(* IEC 61131-3 sources: taksa-factory-simulator/sample_programs, 16 files *)

(* ---- CNCMachiningPLC10.st ---- *)
PROGRAM PLC10_CNC

VAR
    cycle_time : REAL := 120.0;
    throughput : REAL := 30.0;

    dimension_ok : BOOL := TRUE;
    surface_finish : REAL := 0.95;

    tool_break_alarm : BOOL := FALSE;

    spindle_energy : REAL := 50.0;

    machine_idle : REAL := 0.0;

    spindle_load : REAL := 70.0;
    tool_life : REAL := 100.0;

    rand : REAL;
    tick : DINT;
END_VAR

VAR_EXTERNAL
    reg_cycle_time_x10 : UINT;
    reg_throughput_x10 : UINT;
    reg_dimension_ok : UINT;
    reg_surface_finish_x1000 : UINT;
    reg_tool_break_alarm : UINT;
    reg_spindle_energy_x10 : UINT;
    reg_machine_idle_x10 : UINT;
    reg_spindle_load_x10 : UINT;
    reg_tool_life_x10 : UINT;
END_VAR

rand := DINT_TO_REAL((tick * 41) MOD 100) / 100.0;
tick := tick + 1;

cycle_time := 100.0 + (rand * 40.0);
throughput := 3600.0 / cycle_time;

spindle_load := 60.0 + (rand * 30.0);

IF rand < 0.01 THEN
    tool_break_alarm := TRUE;
    dimension_ok := FALSE;
END_IF;

tool_life := tool_life - 0.001;

spindle_energy := spindle_load * 0.8;

(* Export live values to Modbus holding registers %MW0.. *)
reg_cycle_time_x10 := REAL_TO_UINT(cycle_time * 10.0);
reg_throughput_x10 := REAL_TO_UINT(throughput * 10.0);
IF dimension_ok THEN
    reg_dimension_ok := 1;
ELSE
    reg_dimension_ok := 0;
END_IF;
reg_surface_finish_x1000 := REAL_TO_UINT(surface_finish * 1000.0);
IF tool_break_alarm THEN
    reg_tool_break_alarm := 1;
ELSE
    reg_tool_break_alarm := 0;
END_IF;
reg_spindle_energy_x10 := REAL_TO_UINT(spindle_energy * 10.0);
reg_machine_idle_x10 := REAL_TO_UINT(machine_idle * 10.0);
reg_spindle_load_x10 := REAL_TO_UINT(spindle_load * 10.0);
reg_tool_life_x10 := REAL_TO_UINT(tool_life * 10.0);

END_PROGRAM

CONFIGURATION Config0
  RESOURCE Res0 ON PLC
    VAR_GLOBAL
      reg_cycle_time_x10 AT %MW0 : UINT;
      reg_throughput_x10 AT %MW1 : UINT;
      reg_dimension_ok AT %MW2 : UINT;
      reg_surface_finish_x1000 AT %MW3 : UINT;
      reg_tool_break_alarm AT %MW4 : UINT;
      reg_spindle_energy_x10 AT %MW5 : UINT;
      reg_machine_idle_x10 AT %MW6 : UINT;
      reg_spindle_load_x10 AT %MW7 : UINT;
      reg_tool_life_x10 AT %MW8 : UINT;
    END_VAR

    TASK Main(INTERVAL := T#20ms, PRIORITY := 0);
    PROGRAM Inst0 WITH Main : PLC10_CNC;
  END_RESOURCE
END_CONFIGURATION

(* ---- CNCMachiningPLC8.st ---- *)
PROGRAM PLC8_CNC

VAR
    cycle_time : REAL := 120.0;
    throughput : REAL := 30.0;

    dimension_ok : BOOL := TRUE;
    surface_finish : REAL := 0.95;

    tool_break_alarm : BOOL := FALSE;

    spindle_energy : REAL := 50.0;

    machine_idle : REAL := 0.0;

    spindle_load : REAL := 70.0;
    tool_life : REAL := 100.0;

    rand : REAL;
    tick : DINT;
END_VAR

VAR_EXTERNAL
    reg_cycle_time_x10 : UINT;
    reg_throughput_x10 : UINT;
    reg_dimension_ok : UINT;
    reg_surface_finish_x1000 : UINT;
    reg_tool_break_alarm : UINT;
    reg_spindle_energy_x10 : UINT;
    reg_machine_idle_x10 : UINT;
    reg_spindle_load_x10 : UINT;
    reg_tool_life_x10 : UINT;
END_VAR

rand := DINT_TO_REAL((tick * 41) MOD 100) / 100.0;
tick := tick + 1;

cycle_time := 100.0 + (rand * 40.0);
throughput := 3600.0 / cycle_time;

spindle_load := 60.0 + (rand * 30.0);

IF rand < 0.01 THEN
    tool_break_alarm := TRUE;
    dimension_ok := FALSE;
END_IF;

tool_life := tool_life - 0.001;

spindle_energy := spindle_load * 0.8;

(* Export live values to Modbus holding registers %MW0.. *)
reg_cycle_time_x10 := REAL_TO_UINT(cycle_time * 10.0);
reg_throughput_x10 := REAL_TO_UINT(throughput * 10.0);
IF dimension_ok THEN
    reg_dimension_ok := 1;
ELSE
    reg_dimension_ok := 0;
END_IF;
reg_surface_finish_x1000 := REAL_TO_UINT(surface_finish * 1000.0);
IF tool_break_alarm THEN
    reg_tool_break_alarm := 1;
ELSE
    reg_tool_break_alarm := 0;
END_IF;
reg_spindle_energy_x10 := REAL_TO_UINT(spindle_energy * 10.0);
reg_machine_idle_x10 := REAL_TO_UINT(machine_idle * 10.0);
reg_spindle_load_x10 := REAL_TO_UINT(spindle_load * 10.0);
reg_tool_life_x10 := REAL_TO_UINT(tool_life * 10.0);

END_PROGRAM

CONFIGURATION Config0
  RESOURCE Res0 ON PLC
    VAR_GLOBAL
      reg_cycle_time_x10 AT %MW0 : UINT;
      reg_throughput_x10 AT %MW1 : UINT;
      reg_dimension_ok AT %MW2 : UINT;
      reg_surface_finish_x1000 AT %MW3 : UINT;
      reg_tool_break_alarm AT %MW4 : UINT;
      reg_spindle_energy_x10 AT %MW5 : UINT;
      reg_machine_idle_x10 AT %MW6 : UINT;
      reg_spindle_load_x10 AT %MW7 : UINT;
      reg_tool_life_x10 AT %MW8 : UINT;
    END_VAR

    TASK Main(INTERVAL := T#20ms, PRIORITY := 0);
    PROGRAM Inst0 WITH Main : PLC8_CNC;
  END_RESOURCE
END_CONFIGURATION

(* ---- CNCMachiningPLC9.st ---- *)
PROGRAM PLC9_CNC

VAR
    cycle_time : REAL := 120.0;
    throughput : REAL := 30.0;

    dimension_ok : BOOL := TRUE;
    surface_finish : REAL := 0.95;

    tool_break_alarm : BOOL := FALSE;

    spindle_energy : REAL := 50.0;

    machine_idle : REAL := 0.0;

    spindle_load : REAL := 70.0;
    tool_life : REAL := 100.0;

    rand : REAL;
    tick : DINT;
END_VAR

VAR_EXTERNAL
    reg_cycle_time_x10 : UINT;
    reg_throughput_x10 : UINT;
    reg_dimension_ok : UINT;
    reg_surface_finish_x1000 : UINT;
    reg_tool_break_alarm : UINT;
    reg_spindle_energy_x10 : UINT;
    reg_machine_idle_x10 : UINT;
    reg_spindle_load_x10 : UINT;
    reg_tool_life_x10 : UINT;
END_VAR

rand := DINT_TO_REAL((tick * 41) MOD 100) / 100.0;
tick := tick + 1;

cycle_time := 100.0 + (rand * 40.0);
throughput := 3600.0 / cycle_time;

spindle_load := 60.0 + (rand * 30.0);

IF rand < 0.01 THEN
    tool_break_alarm := TRUE;
    dimension_ok := FALSE;
END_IF;

tool_life := tool_life - 0.001;

spindle_energy := spindle_load * 0.8;

(* Export live values to Modbus holding registers %MW0.. *)
reg_cycle_time_x10 := REAL_TO_UINT(cycle_time * 10.0);
reg_throughput_x10 := REAL_TO_UINT(throughput * 10.0);
IF dimension_ok THEN
    reg_dimension_ok := 1;
ELSE
    reg_dimension_ok := 0;
END_IF;
reg_surface_finish_x1000 := REAL_TO_UINT(surface_finish * 1000.0);
IF tool_break_alarm THEN
    reg_tool_break_alarm := 1;
ELSE
    reg_tool_break_alarm := 0;
END_IF;
reg_spindle_energy_x10 := REAL_TO_UINT(spindle_energy * 10.0);
reg_machine_idle_x10 := REAL_TO_UINT(machine_idle * 10.0);
reg_spindle_load_x10 := REAL_TO_UINT(spindle_load * 10.0);
reg_tool_life_x10 := REAL_TO_UINT(tool_life * 10.0);

END_PROGRAM

CONFIGURATION Config0
  RESOURCE Res0 ON PLC
    VAR_GLOBAL
      reg_cycle_time_x10 AT %MW0 : UINT;
      reg_throughput_x10 AT %MW1 : UINT;
      reg_dimension_ok AT %MW2 : UINT;
      reg_surface_finish_x1000 AT %MW3 : UINT;
      reg_tool_break_alarm AT %MW4 : UINT;
      reg_spindle_energy_x10 AT %MW5 : UINT;
      reg_machine_idle_x10 AT %MW6 : UINT;
      reg_spindle_load_x10 AT %MW7 : UINT;
      reg_tool_life_x10 AT %MW8 : UINT;
    END_VAR

    TASK Main(INTERVAL := T#20ms, PRIORITY := 0);
    PROGRAM Inst0 WITH Main : PLC9_CNC;
  END_RESOURCE
END_CONFIGURATION

(* ---- Cooling.st ---- *)
PROGRAM PLC5_COOLING

VAR
    cooling_time : REAL := 120.0;

    cooling_uniformity : REAL := 0.95;

    temp_alarm : BOOL := FALSE;

    water_usage : REAL := 50.0;

    blockage_time : REAL := 0.0;

    pump_health : REAL := 100.0;

    rand : REAL;
    tick : DINT;
END_VAR

VAR_EXTERNAL
    reg_cooling_time_x10 : UINT;
    reg_cooling_uniformity_x1000 : UINT;
    reg_temp_alarm : UINT;
    reg_water_usage_x10 : UINT;
    reg_blockage_time_x10 : UINT;
    reg_pump_health_x10 : UINT;
END_VAR

rand := DINT_TO_REAL((tick * 29) MOD 100) / 100.0;
tick := tick + 1;

cooling_time := 100.0 + (rand * 40.0);
cooling_uniformity := 0.9 + (rand * 0.1);

IF rand < 0.01 THEN
    temp_alarm := TRUE;
END_IF;

water_usage := 40.0 + (rand * 20.0);

pump_health := pump_health - 0.0003;

(* Export live values to Modbus holding registers %MW0.. *)
reg_cooling_time_x10 := REAL_TO_UINT(cooling_time * 10.0);
reg_cooling_uniformity_x1000 := REAL_TO_UINT(cooling_uniformity * 1000.0);
IF temp_alarm THEN
    reg_temp_alarm := 1;
ELSE
    reg_temp_alarm := 0;
END_IF;
reg_water_usage_x10 := REAL_TO_UINT(water_usage * 10.0);
reg_blockage_time_x10 := REAL_TO_UINT(blockage_time * 10.0);
reg_pump_health_x10 := REAL_TO_UINT(pump_health * 10.0);

END_PROGRAM

CONFIGURATION Config0
  RESOURCE Res0 ON PLC
    VAR_GLOBAL
      reg_cooling_time_x10 AT %MW0 : UINT;
      reg_cooling_uniformity_x1000 AT %MW1 : UINT;
      reg_temp_alarm AT %MW2 : UINT;
      reg_water_usage_x10 AT %MW3 : UINT;
      reg_blockage_time_x10 AT %MW4 : UINT;
      reg_pump_health_x10 AT %MW5 : UINT;
    END_VAR

    TASK Main(INTERVAL := T#20ms, PRIORITY := 0);
    PROGRAM Inst0 WITH Main : PLC5_COOLING;
  END_RESOURCE
END_CONFIGURATION

(* ---- Degassing.st ---- *)
PROGRAM PLC3_DEGASS

VAR
    treatment_cycle_time : REAL := 60.0;

    gas_content_level : REAL := 0.02;

    gas_leak_alarm : BOOL := FALSE;

    gas_consumption : REAL := 10.0;

    idle_time : REAL := 0.0;

    rotor_health : REAL := 100.0;

    rand : REAL;
    tick : DINT;
END_VAR

VAR_EXTERNAL
    reg_treatment_cycle_time_x10 : UINT;
    reg_gas_content_level_x10000 : UINT;
    reg_gas_leak_alarm : UINT;
    reg_gas_consumption_x10 : UINT;
    reg_idle_time_x10 : UINT;
    reg_rotor_health_x10 : UINT;
END_VAR

rand := DINT_TO_REAL((tick * 19) MOD 100) / 100.0;
tick := tick + 1;

gas_content_level := 0.01 + (rand * 0.02);

IF rand < 0.005 THEN
    gas_leak_alarm := TRUE;
ELSE
    gas_leak_alarm := FALSE;
END_IF;

gas_consumption := 8.0 + (rand * 4.0);

rotor_health := rotor_health - 0.0004;

(* Export live values to Modbus holding registers %MW0.. *)
reg_treatment_cycle_time_x10 := REAL_TO_UINT(treatment_cycle_time * 10.0);
reg_gas_content_level_x10000 := REAL_TO_UINT(gas_content_level * 10000.0);
IF gas_leak_alarm THEN
    reg_gas_leak_alarm := 1;
ELSE
    reg_gas_leak_alarm := 0;
END_IF;
reg_gas_consumption_x10 := REAL_TO_UINT(gas_consumption * 10.0);
reg_idle_time_x10 := REAL_TO_UINT(idle_time * 10.0);
reg_rotor_health_x10 := REAL_TO_UINT(rotor_health * 10.0);

END_PROGRAM

CONFIGURATION Config0
  RESOURCE Res0 ON PLC
    VAR_GLOBAL
      reg_treatment_cycle_time_x10 AT %MW0 : UINT;
      reg_gas_content_level_x10000 AT %MW1 : UINT;
      reg_gas_leak_alarm AT %MW2 : UINT;
      reg_gas_consumption_x10 AT %MW3 : UINT;
      reg_idle_time_x10 AT %MW4 : UINT;
      reg_rotor_health_x10 AT %MW5 : UINT;
    END_VAR

    TASK Main(INTERVAL := T#20ms, PRIORITY := 0);
    PROGRAM Inst0 WITH Main : PLC3_DEGASS;
  END_RESOURCE
END_CONFIGURATION

(* ---- FinalInspection.st ---- *)
PROGRAM PLC13_FINAL_INSPECTION

VAR
    inspection_cycle : REAL := 30.0;

    crack_detected : BOOL := FALSE;
    pass_fail : BOOL := TRUE;

    radiation_alarm : BOOL := FALSE;

    energy_usage : REAL := 50.0;

    reinspection_time : REAL := 0.0;

    sensor_health : REAL := 100.0;

    rand : REAL;
    tick : DINT;
END_VAR

VAR_EXTERNAL
    reg_inspection_cycle_x10 : UINT;
    reg_crack_detected : UINT;
    reg_pass_fail : UINT;
    reg_radiation_alarm : UINT;
    reg_energy_usage_x10 : UINT;
    reg_reinspection_time_x10 : UINT;
    reg_sensor_health_x10 : UINT;
END_VAR

rand := DINT_TO_REAL((tick * 53) MOD 100) / 100.0;
tick := tick + 1;

IF rand < 0.01 THEN
    crack_detected := TRUE;
    pass_fail := FALSE;
END_IF;

sensor_health := sensor_health - 0.0002;

(* Export live values to Modbus holding registers %MW0.. *)
reg_inspection_cycle_x10 := REAL_TO_UINT(inspection_cycle * 10.0);
IF crack_detected THEN
    reg_crack_detected := 1;
ELSE
    reg_crack_detected := 0;
END_IF;
IF pass_fail THEN
    reg_pass_fail := 1;
ELSE
    reg_pass_fail := 0;
END_IF;
IF radiation_alarm THEN
    reg_radiation_alarm := 1;
ELSE
    reg_radiation_alarm := 0;
END_IF;
reg_energy_usage_x10 := REAL_TO_UINT(energy_usage * 10.0);
reg_reinspection_time_x10 := REAL_TO_UINT(reinspection_time * 10.0);
reg_sensor_health_x10 := REAL_TO_UINT(sensor_health * 10.0);

END_PROGRAM

CONFIGURATION Config0
  RESOURCE Res0 ON PLC
    VAR_GLOBAL
      reg_inspection_cycle_x10 AT %MW0 : UINT;
      reg_crack_detected AT %MW1 : UINT;
      reg_pass_fail AT %MW2 : UINT;
      reg_radiation_alarm AT %MW3 : UINT;
      reg_energy_usage_x10 AT %MW4 : UINT;
      reg_reinspection_time_x10 AT %MW5 : UINT;
      reg_sensor_health_x10 AT %MW6 : UINT;
    END_VAR

    TASK Main(INTERVAL := T#20ms, PRIORITY := 0);
    PROGRAM Inst0 WITH Main : PLC13_FINAL_INSPECTION;
  END_RESOURCE
END_CONFIGURATION

(* ---- HeatTreatment.st ---- *)
PROGRAM PLC6_HEATTREAT

VAR
    batch_cycle_time : REAL := 3600.0;

    hardness : REAL := 80.0;
    temperature_profile : REAL := 500.0;

    furnace_alarm : BOOL := FALSE;

    fuel_consumption : REAL := 300.0;

    downtime : REAL := 0.0;

    heater_health : REAL := 100.0;

    rand : REAL;
    tick : DINT;
END_VAR

VAR_EXTERNAL
    reg_batch_cycle_time_s : UINT;
    reg_hardness_x10 : UINT;
    reg_temperature_profile_x10 : UINT;
    reg_furnace_alarm : UINT;
    reg_fuel_consumption_x10 : UINT;
    reg_downtime_x10 : UINT;
    reg_heater_health_x10 : UINT;
END_VAR

rand := DINT_TO_REAL((tick * 31) MOD 100) / 100.0;
tick := tick + 1;

temperature_profile := 480.0 + (rand * 40.0);

IF rand < 0.01 THEN
    furnace_alarm := TRUE;
END_IF;

fuel_consumption := 250.0 + (rand * 100.0);

heater_health := heater_health - 0.0004;

(* Export live values to Modbus holding registers %MW0.. *)
reg_batch_cycle_time_s := REAL_TO_UINT(batch_cycle_time);
reg_hardness_x10 := REAL_TO_UINT(hardness * 10.0);
reg_temperature_profile_x10 := REAL_TO_UINT(temperature_profile * 10.0);
IF furnace_alarm THEN
    reg_furnace_alarm := 1;
ELSE
    reg_furnace_alarm := 0;
END_IF;
reg_fuel_consumption_x10 := REAL_TO_UINT(fuel_consumption * 10.0);
reg_downtime_x10 := REAL_TO_UINT(downtime * 10.0);
reg_heater_health_x10 := REAL_TO_UINT(heater_health * 10.0);

END_PROGRAM

CONFIGURATION Config0
  RESOURCE Res0 ON PLC
    VAR_GLOBAL
      reg_batch_cycle_time_s AT %MW0 : UINT;
      reg_hardness_x10 AT %MW1 : UINT;
      reg_temperature_profile_x10 AT %MW2 : UINT;
      reg_furnace_alarm AT %MW3 : UINT;
      reg_fuel_consumption_x10 AT %MW4 : UINT;
      reg_downtime_x10 AT %MW5 : UINT;
      reg_heater_health_x10 AT %MW6 : UINT;
    END_VAR

    TASK Main(INTERVAL := T#20ms, PRIORITY := 0);
    PROGRAM Inst0 WITH Main : PLC6_HEATTREAT;
  END_RESOURCE
END_CONFIGURATION

(* ---- Inspection.st ---- *)
PROGRAM PLC11_INSPECTION

VAR
    inspection_rate : REAL := 60.0;

    defect_detected : BOOL := FALSE;
    defect_type : INT := 0;

    camera_fault : BOOL := FALSE;

    system_energy : REAL := 20.0;

    inspection_delay : REAL := 0.0;

    camera_health : REAL := 100.0;

    rand : REAL;
    tick : DINT;
END_VAR

VAR_EXTERNAL
    reg_inspection_rate_x10 : UINT;
    reg_defect_detected : UINT;
    reg_defect_type : UINT;
    reg_camera_fault : UINT;
    reg_system_energy_x10 : UINT;
    reg_inspection_delay_x10 : UINT;
    reg_camera_health_x10 : UINT;
END_VAR

rand := DINT_TO_REAL((tick * 43) MOD 100) / 100.0;
tick := tick + 1;

IF rand < 0.02 THEN
    defect_detected := TRUE;
    defect_type := 1;
END_IF;

IF rand < 0.005 THEN
    camera_fault := TRUE;
END_IF;

camera_health := camera_health - 0.0002;

(* Export live values to Modbus holding registers %MW0.. *)
reg_inspection_rate_x10 := REAL_TO_UINT(inspection_rate * 10.0);
IF defect_detected THEN
    reg_defect_detected := 1;
ELSE
    reg_defect_detected := 0;
END_IF;
IF defect_type < 0 THEN
    reg_defect_type := 0;
ELSE
    reg_defect_type := INT_TO_UINT(defect_type);
END_IF;
IF camera_fault THEN
    reg_camera_fault := 1;
ELSE
    reg_camera_fault := 0;
END_IF;
reg_system_energy_x10 := REAL_TO_UINT(system_energy * 10.0);
reg_inspection_delay_x10 := REAL_TO_UINT(inspection_delay * 10.0);
reg_camera_health_x10 := REAL_TO_UINT(camera_health * 10.0);

END_PROGRAM

CONFIGURATION Config0
  RESOURCE Res0 ON PLC
    VAR_GLOBAL
      reg_inspection_rate_x10 AT %MW0 : UINT;
      reg_defect_detected AT %MW1 : UINT;
      reg_defect_type AT %MW2 : UINT;
      reg_camera_fault AT %MW3 : UINT;
      reg_system_energy_x10 AT %MW4 : UINT;
      reg_inspection_delay_x10 AT %MW5 : UINT;
      reg_camera_health_x10 AT %MW6 : UINT;
    END_VAR

    TASK Main(INTERVAL := T#20ms, PRIORITY := 0);
    PROGRAM Inst0 WITH Main : PLC11_INSPECTION;
  END_RESOURCE
END_CONFIGURATION

(* ---- MeltingFurnace.st ---- *)
PROGRAM PLC2_FURNACE

VAR
    melt_rate : REAL := 100.0;
    tap_time  : REAL := 0.0;

    metal_temperature : REAL := 700.0;
    composition : REAL := 0.95;

    overheat_alarm : BOOL := FALSE;

    energy_consumption : REAL := 500.0;

    furnace_downtime : REAL := 0.0;

    refractory_health : REAL := 100.0;

    rand : REAL;
    tick : DINT;
END_VAR

VAR_EXTERNAL
    reg_melt_rate_x10 : UINT;
    reg_tap_time_x10 : UINT;
    reg_metal_temperature_x10 : UINT;
    reg_composition_x1000 : UINT;
    reg_overheat_alarm : UINT;
    reg_energy_consumption_x10 : UINT;
    reg_furnace_downtime_x10 : UINT;
    reg_refractory_health_x10 : UINT;
END_VAR

rand := DINT_TO_REAL((tick * 17) MOD 100) / 100.0;
tick := tick + 1;

metal_temperature := 680.0 + (rand * 50.0);

IF metal_temperature > 720.0 THEN
    overheat_alarm := TRUE;
    furnace_downtime := furnace_downtime + 0.1;
ELSE
    overheat_alarm := FALSE;
END_IF;

melt_rate := 90.0 + (rand * 20.0);
energy_consumption := melt_rate * 4.0;

refractory_health := refractory_health - 0.0003;

tap_time := tap_time + 0.1;

(* Export live values to Modbus holding registers %MW0.. *)
reg_melt_rate_x10 := REAL_TO_UINT(melt_rate * 10.0);
reg_tap_time_x10 := REAL_TO_UINT(tap_time * 10.0);
reg_metal_temperature_x10 := REAL_TO_UINT(metal_temperature * 10.0);
reg_composition_x1000 := REAL_TO_UINT(composition * 1000.0);
IF overheat_alarm THEN
    reg_overheat_alarm := 1;
ELSE
    reg_overheat_alarm := 0;
END_IF;
reg_energy_consumption_x10 := REAL_TO_UINT(energy_consumption * 10.0);
reg_furnace_downtime_x10 := REAL_TO_UINT(furnace_downtime * 10.0);
reg_refractory_health_x10 := REAL_TO_UINT(refractory_health * 10.0);

END_PROGRAM

CONFIGURATION Config0
  RESOURCE Res0 ON PLC
    VAR_GLOBAL
      reg_melt_rate_x10 AT %MW0 : UINT;
      reg_tap_time_x10 AT %MW1 : UINT;
      reg_metal_temperature_x10 AT %MW2 : UINT;
      reg_composition_x1000 AT %MW3 : UINT;
      reg_overheat_alarm AT %MW4 : UINT;
      reg_energy_consumption_x10 AT %MW5 : UINT;
      reg_furnace_downtime_x10 AT %MW6 : UINT;
      reg_refractory_health_x10 AT %MW7 : UINT;
    END_VAR

    TASK Main(INTERVAL := T#20ms, PRIORITY := 0);
    PROGRAM Inst0 WITH Main : PLC2_FURNACE;
  END_RESOURCE
END_CONFIGURATION

(* ---- Packing.st ---- *)
PROGRAM PLC14_PACKING

VAR
    packing_rate : REAL := 100.0;

    packing_ok : BOOL := TRUE;

    jam_alarm : BOOL := FALSE;

    material_usage : REAL := 20.0;

    downtime : REAL := 0.0;

    robot_health : REAL := 100.0;

    rand : REAL;
    tick : DINT;
END_VAR

VAR_EXTERNAL
    reg_packing_rate_x10 : UINT;
    reg_packing_ok : UINT;
    reg_jam_alarm : UINT;
    reg_material_usage_x10 : UINT;
    reg_downtime_x10 : UINT;
    reg_robot_health_x10 : UINT;
END_VAR

rand := DINT_TO_REAL((tick * 59) MOD 100) / 100.0;
tick := tick + 1;

IF rand < 0.01 THEN
    jam_alarm := TRUE;
END_IF;

robot_health := robot_health - 0.0003;

(* Export live values to Modbus holding registers %MW0.. *)
reg_packing_rate_x10 := REAL_TO_UINT(packing_rate * 10.0);
IF packing_ok THEN
    reg_packing_ok := 1;
ELSE
    reg_packing_ok := 0;
END_IF;
IF jam_alarm THEN
    reg_jam_alarm := 1;
ELSE
    reg_jam_alarm := 0;
END_IF;
reg_material_usage_x10 := REAL_TO_UINT(material_usage * 10.0);
reg_downtime_x10 := REAL_TO_UINT(downtime * 10.0);
reg_robot_health_x10 := REAL_TO_UINT(robot_health * 10.0);

END_PROGRAM

CONFIGURATION Config0
  RESOURCE Res0 ON PLC
    VAR_GLOBAL
      reg_packing_rate_x10 AT %MW0 : UINT;
      reg_packing_ok AT %MW1 : UINT;
      reg_jam_alarm AT %MW2 : UINT;
      reg_material_usage_x10 AT %MW3 : UINT;
      reg_downtime_x10 AT %MW4 : UINT;
      reg_robot_health_x10 AT %MW5 : UINT;
    END_VAR

    TASK Main(INTERVAL := T#20ms, PRIORITY := 0);
    PROGRAM Inst0 WITH Main : PLC14_PACKING;
  END_RESOURCE
END_CONFIGURATION

(* ---- Painting.st ---- *)
PROGRAM PLC12_PAINT

VAR
    coating_rate : REAL := 40.0;

    thickness : REAL := 50.0;
    finish_quality : REAL := 0.95;

    oven_alarm : BOOL := FALSE;

    powder_usage : REAL := 10.0;
    energy : REAL := 200.0;

    line_stop_time : REAL := 0.0;

    nozzle_health : REAL := 100.0;

    rand : REAL;
    tick : DINT;
END_VAR

VAR_EXTERNAL
    reg_coating_rate_x10 : UINT;
    reg_thickness_x10 : UINT;
    reg_finish_quality_x1000 : UINT;
    reg_oven_alarm : UINT;
    reg_powder_usage_x10 : UINT;
    reg_energy_x10 : UINT;
    reg_line_stop_time_x10 : UINT;
    reg_nozzle_health_x10 : UINT;
END_VAR

rand := DINT_TO_REAL((tick * 47) MOD 100) / 100.0;
tick := tick + 1;

thickness := 45.0 + (rand * 10.0);

IF rand < 0.01 THEN
    oven_alarm := TRUE;
END_IF;

nozzle_health := nozzle_health - 0.0003;

(* Export live values to Modbus holding registers %MW0.. *)
reg_coating_rate_x10 := REAL_TO_UINT(coating_rate * 10.0);
reg_thickness_x10 := REAL_TO_UINT(thickness * 10.0);
reg_finish_quality_x1000 := REAL_TO_UINT(finish_quality * 1000.0);
IF oven_alarm THEN
    reg_oven_alarm := 1;
ELSE
    reg_oven_alarm := 0;
END_IF;
reg_powder_usage_x10 := REAL_TO_UINT(powder_usage * 10.0);
reg_energy_x10 := REAL_TO_UINT(energy * 10.0);
reg_line_stop_time_x10 := REAL_TO_UINT(line_stop_time * 10.0);
reg_nozzle_health_x10 := REAL_TO_UINT(nozzle_health * 10.0);

END_PROGRAM

CONFIGURATION Config0
  RESOURCE Res0 ON PLC
    VAR_GLOBAL
      reg_coating_rate_x10 AT %MW0 : UINT;
      reg_thickness_x10 AT %MW1 : UINT;
      reg_finish_quality_x1000 AT %MW2 : UINT;
      reg_oven_alarm AT %MW3 : UINT;
      reg_powder_usage_x10 AT %MW4 : UINT;
      reg_energy_x10 AT %MW5 : UINT;
      reg_line_stop_time_x10 AT %MW6 : UINT;
      reg_nozzle_health_x10 AT %MW7 : UINT;
    END_VAR

    TASK Main(INTERVAL := T#20ms, PRIORITY := 0);
    PROGRAM Inst0 WITH Main : PLC12_PAINT;
  END_RESOURCE
END_CONFIGURATION

(* ---- Press.st ---- *)
PROGRAM PLC4_PRESS

VAR
    cycle_time : REAL := 30.0;
    parts_per_hour : REAL := 100.0;

    porosity_flag : BOOL := FALSE;
    fill_quality : REAL := 0.95;

    pressure_alarm : BOOL := FALSE;

    hydraulic_energy : REAL := 200.0;

    press_idle_time : REAL := 0.0;

    press_load : REAL := 70.0;
    die_health : REAL := 100.0;

    rand : REAL;
    tick : DINT;
END_VAR

VAR_EXTERNAL
    reg_cycle_time_x10 : UINT;
    reg_parts_per_hour_x10 : UINT;
    reg_porosity_flag : UINT;
    reg_fill_quality_x1000 : UINT;
    reg_pressure_alarm : UINT;
    reg_hydraulic_energy_x10 : UINT;
    reg_press_idle_time_x10 : UINT;
    reg_press_load_x10 : UINT;
    reg_die_health_x10 : UINT;
END_VAR

rand := DINT_TO_REAL((tick * 23) MOD 100) / 100.0;
tick := tick + 1;

cycle_time := 25.0 + (rand * 10.0);
parts_per_hour := 3600.0 / cycle_time;

fill_quality := 0.9 + (rand * 0.1);

IF rand < 0.02 THEN
    porosity_flag := TRUE;
END_IF;

press_load := 60.0 + (rand * 30.0);

IF press_load > 85.0 THEN
    pressure_alarm := TRUE;
END_IF;

hydraulic_energy := press_load * 2.5;

die_health := die_health - 0.0005;

(* Export live values to Modbus holding registers %MW0.. *)
reg_cycle_time_x10 := REAL_TO_UINT(cycle_time * 10.0);
reg_parts_per_hour_x10 := REAL_TO_UINT(parts_per_hour * 10.0);
IF porosity_flag THEN
    reg_porosity_flag := 1;
ELSE
    reg_porosity_flag := 0;
END_IF;
reg_fill_quality_x1000 := REAL_TO_UINT(fill_quality * 1000.0);
IF pressure_alarm THEN
    reg_pressure_alarm := 1;
ELSE
    reg_pressure_alarm := 0;
END_IF;
reg_hydraulic_energy_x10 := REAL_TO_UINT(hydraulic_energy * 10.0);
reg_press_idle_time_x10 := REAL_TO_UINT(press_idle_time * 10.0);
reg_press_load_x10 := REAL_TO_UINT(press_load * 10.0);
reg_die_health_x10 := REAL_TO_UINT(die_health * 10.0);

END_PROGRAM

CONFIGURATION Config0
  RESOURCE Res0 ON PLC
    VAR_GLOBAL
      reg_cycle_time_x10 AT %MW0 : UINT;
      reg_parts_per_hour_x10 AT %MW1 : UINT;
      reg_porosity_flag AT %MW2 : UINT;
      reg_fill_quality_x1000 AT %MW3 : UINT;
      reg_pressure_alarm AT %MW4 : UINT;
      reg_hydraulic_energy_x10 AT %MW5 : UINT;
      reg_press_idle_time_x10 AT %MW6 : UINT;
      reg_press_load_x10 AT %MW7 : UINT;
      reg_die_health_x10 AT %MW8 : UINT;
    END_VAR

    TASK Main(INTERVAL := T#20ms, PRIORITY := 0);
    PROGRAM Inst0 WITH Main : PLC4_PRESS;
  END_RESOURCE
END_CONFIGURATION

(* ---- program.st ---- *)
PROGRAM main
VAR
    start_button AT %IX0.0 : BOOL;
    motor        AT %QX0.0 : BOOL;
    counter      AT %MW0   : INT := 0;
END_VAR

(* Logic *)
IF start_button THEN
    motor := TRUE;
    counter := counter + 1;
ELSE
    motor := FALSE;
END_IF;

END_PROGRAM

(* ---- RawMaterialHandling.st ---- *)
PROGRAM PLC1_RAW_MATERIAL

VAR

    material_feed_rate : REAL := 50.0;
    material_available : BOOL := TRUE;

    material_composition_ok : BOOL := TRUE;

    overload_alarm : BOOL := FALSE;

    energy_usage_conveyor : REAL := 5.0;

    feeder_idle_time : REAL := 0.0;

    motor_health : REAL := 100.0;

    rand : REAL := 0.5;
    tick : DINT := 0;
END_VAR

VAR_EXTERNAL
    reg_material_feed_rate_x10 : UINT;
    reg_material_available : UINT;
    reg_material_composition_ok : UINT;
    reg_overload_alarm : UINT;
    reg_energy_usage_conveyor_x10 : UINT;
    reg_feeder_idle_time_x10 : UINT;
    reg_motor_health_x10 : UINT;
END_VAR

rand := DINT_TO_REAL((tick * 13) MOD 100) / 100.0;
tick := tick + 1;

material_feed_rate := 45.0 + (rand * 10.0);

IF rand < 0.01 THEN
    overload_alarm := TRUE;
ELSE
    overload_alarm := FALSE;
END_IF;

IF NOT material_available THEN
    feeder_idle_time := feeder_idle_time + 0.1;
END_IF;

motor_health := motor_health - 0.0005;

energy_usage_conveyor := material_feed_rate * 0.1;

(* Export live values to Modbus holding registers %MW0.. *)
reg_material_feed_rate_x10 := REAL_TO_UINT(material_feed_rate * 10.0);
IF material_available THEN
    reg_material_available := 1;
ELSE
    reg_material_available := 0;
END_IF;
IF material_composition_ok THEN
    reg_material_composition_ok := 1;
ELSE
    reg_material_composition_ok := 0;
END_IF;
IF overload_alarm THEN
    reg_overload_alarm := 1;
ELSE
    reg_overload_alarm := 0;
END_IF;
reg_energy_usage_conveyor_x10 := REAL_TO_UINT(energy_usage_conveyor * 10.0);
reg_feeder_idle_time_x10 := REAL_TO_UINT(feeder_idle_time * 10.0);
reg_motor_health_x10 := REAL_TO_UINT(motor_health * 10.0);

END_PROGRAM

CONFIGURATION Config0
  RESOURCE Res0 ON PLC
    VAR_GLOBAL
      reg_material_feed_rate_x10 AT %MW0 : UINT;
      reg_material_available AT %MW1 : UINT;
      reg_material_composition_ok AT %MW2 : UINT;
      reg_overload_alarm AT %MW3 : UINT;
      reg_energy_usage_conveyor_x10 AT %MW4 : UINT;
      reg_feeder_idle_time_x10 AT %MW5 : UINT;
      reg_motor_health_x10 AT %MW6 : UINT;
    END_VAR

    TASK Main(INTERVAL := T#20ms, PRIORITY := 0);
    PROGRAM Inst0 WITH Main : PLC1_RAW_MATERIAL;
  END_RESOURCE
END_CONFIGURATION

(* ---- ShotBlasting.st ---- *)
PROGRAM PLC7_SHOTBLAST

VAR
    cycle_time : REAL := 60.0;

    surface_cleanliness : REAL := 0.95;

    vibration_alarm : BOOL := FALSE;

    media_usage : REAL := 5.0;

    jam_time : REAL := 0.0;

    turbine_health : REAL := 100.0;

    rand : REAL;
    tick : DINT;
END_VAR

VAR_EXTERNAL
    reg_cycle_time_x10 : UINT;
    reg_surface_cleanliness_x1000 : UINT;
    reg_vibration_alarm : UINT;
    reg_media_usage_x10 : UINT;
    reg_jam_time_x10 : UINT;
    reg_turbine_health_x10 : UINT;
END_VAR

rand := DINT_TO_REAL((tick * 37) MOD 100) / 100.0;
tick := tick + 1;

surface_cleanliness := 0.9 + (rand * 0.1);

IF rand < 0.01 THEN
    vibration_alarm := TRUE;
END_IF;

media_usage := 4.0 + (rand * 2.0);

turbine_health := turbine_health - 0.0003;

(* Export live values to Modbus holding registers %MW0.. *)
reg_cycle_time_x10 := REAL_TO_UINT(cycle_time * 10.0);
reg_surface_cleanliness_x1000 := REAL_TO_UINT(surface_cleanliness * 1000.0);
IF vibration_alarm THEN
    reg_vibration_alarm := 1;
ELSE
    reg_vibration_alarm := 0;
END_IF;
reg_media_usage_x10 := REAL_TO_UINT(media_usage * 10.0);
reg_jam_time_x10 := REAL_TO_UINT(jam_time * 10.0);
reg_turbine_health_x10 := REAL_TO_UINT(turbine_health * 10.0);

END_PROGRAM

CONFIGURATION Config0
  RESOURCE Res0 ON PLC
    VAR_GLOBAL
      reg_cycle_time_x10 AT %MW0 : UINT;
      reg_surface_cleanliness_x1000 AT %MW1 : UINT;
      reg_vibration_alarm AT %MW2 : UINT;
      reg_media_usage_x10 AT %MW3 : UINT;
      reg_jam_time_x10 AT %MW4 : UINT;
      reg_turbine_health_x10 AT %MW5 : UINT;
    END_VAR

    TASK Main(INTERVAL := T#20ms, PRIORITY := 0);
    PROGRAM Inst0 WITH Main : PLC7_SHOTBLAST;
  END_RESOURCE
END_CONFIGURATION

(* ---- Utilities.st ---- *)
PROGRAM PLC15_UTILS

VAR
    supply_rate : REAL := 100.0;

    pressure_stability : REAL := 0.95;

    power_fault : BOOL := FALSE;

    total_energy : REAL := 1000.0;

    outage_time : REAL := 0.0;

    compressor_health : REAL := 100.0;

    rand : REAL;
    tick : DINT;
END_VAR

VAR_EXTERNAL
    reg_supply_rate_x10 : UINT;
    reg_pressure_stability_x1000 : UINT;
    reg_power_fault : UINT;
    reg_total_energy_x10 : UINT;
    reg_outage_time_x10 : UINT;
    reg_compressor_health_x10 : UINT;
END_VAR

rand := DINT_TO_REAL((tick * 61) MOD 100) / 100.0;
tick := tick + 1;

pressure_stability := 0.9 + (rand * 0.1);

IF rand < 0.005 THEN
    power_fault := TRUE;
    outage_time := outage_time + 0.1;
END_IF;

total_energy := total_energy + (rand * 10.0);

compressor_health := compressor_health - 0.0004;

(* Export live values to Modbus holding registers %MW0.. *)
reg_supply_rate_x10 := REAL_TO_UINT(supply_rate * 10.0);
reg_pressure_stability_x1000 := REAL_TO_UINT(pressure_stability * 1000.0);
IF power_fault THEN
    reg_power_fault := 1;
ELSE
    reg_power_fault := 0;
END_IF;
reg_total_energy_x10 := REAL_TO_UINT(total_energy * 10.0);
reg_outage_time_x10 := REAL_TO_UINT(outage_time * 10.0);
reg_compressor_health_x10 := REAL_TO_UINT(compressor_health * 10.0);

END_PROGRAM

CONFIGURATION Config0
  RESOURCE Res0 ON PLC
    VAR_GLOBAL
      reg_supply_rate_x10 AT %MW0 : UINT;
      reg_pressure_stability_x1000 AT %MW1 : UINT;
      reg_power_fault AT %MW2 : UINT;
      reg_total_energy_x10 AT %MW3 : UINT;
      reg_outage_time_x10 AT %MW4 : UINT;
      reg_compressor_health_x10 AT %MW5 : UINT;
    END_VAR

    TASK Main(INTERVAL := T#20ms, PRIORITY := 0);
    PROGRAM Inst0 WITH Main : PLC15_UTILS;
  END_RESOURCE
END_CONFIGURATION
